ABB RAPID module: RsTempModule.modx

MODULE RsTempModule
PROC RsTempPath()
        SetSysData wobj0;
        SetSysData tool0;
ENDPROC

ENDMODULE
